(* Logix 5000 project; controller MECO9497 vendor 1 type 14 code 106 rev 21.11; software revision 21.00; part 4 of 4 *)
(* tags used below, declared in another part *)
   AAH_200_SP : REAL;
   AAH_200_SP_H : BOOL;
   AAH_200_SP_N : BOOL;
   AAH_200_SP_O : REAL;
   ALERT_ALARM_SU_DELAY : TIMER;
   ALERT_ALARM_SU_DELAY_H : BOOL;
   ALERT_ALARM_SU_DELAY_N : BOOL;
   ALERT_ALARM_SU_DELAY_O : DINT;
   DIST_COND_ALRM_STARTUP_TIME_H : BOOL;
   DIST_COND_ALRM_STARTUP_TIME_N : BOOL;
   DIST_COND_ALRM_STARTUP_TIME_O : REAL;
   DIST_COND_ALRM_STARTUP_TMR : TIMER;
   DIST_PUMP_START_SP : REAL;
   DIST_PUMP_START_SP_H : BOOL;
   DIST_PUMP_START_SP_N : BOOL;
   DIST_PUMP_START_SP_OIT : REAL;
   DIST_PUMP_STOP_SP : REAL;
   DIST_PUMP_STOP_SP_H : BOOL;
   DIST_PUMP_STOP_SP_N : BOOL;
   DIST_PUMP_STOP_SP_OIT : DINT;
   DSTLT_TEMP_ALRM_SU_DELAY : TIMER;
   DSTLT_TEMP_ALRM_SU_DELAY_H : BOOL;
   DSTLT_TEMP_ALRM_SU_DELAY_N : BOOL;
   DSTLT_TEMP_ALRM_SU_DELAY_O : REAL;
   ENGINEER : BOOL;
   EVAP_PRESSURE_PERM_TIME_H : BOOL;
   EVAP_PRESSURE_PERM_TIME_N : BOOL;
   EVAP_PRESSURE_PERM_TIME_O : REAL;
   EVAP_PRESSURE_PERM_TIMER : TIMER;
   EXCESS_DIST_TIME_SP_H : BOOL;
   EXCESS_DIST_TIME_SP_N : BOOL;
   EXCESS_DIST_TIME_SP_OIT : REAL;
   EXCESS_DSTLT_DRAIN_TIMER : TIMER;
   FC_300_SP : DINT;
   FC_300_SP_H : BOOL;
   FC_300_SP_N : BOOL;
   FC_300_SP_O : DINT;
   IAL_100_SP : REAL;
   IAL_100_SP_H : BOOL;
   IAL_100_SP_N : BOOL;
   IAL_100_SP_OIT : REAL;
   LAAH_100_ALERT_H : BOOL;
   LAAH_100_ALERT_N : BOOL;
   LAAH_100_ALERT_O : DINT;
   LAAH_100_SP : DINT;
   LAAL_100_ALERT_H : BOOL;
   LAAL_100_ALERT_N : BOOL;
   LAAL_100_ALERT_O : DINT;
   LAAL_100_SP : DINT;
   LAH_100_SP : REAL;
   LAH_100_SP_H : BOOL;
   LAH_100_SP_N : BOOL;
   LAH_100_SP_OIT : REAL;
   LAL_100_SP : REAL;
   LAL_100_SP_H : BOOL;
   LAL_100_SP_N : BOOL;
   LAL_100_SP_OIT : REAL;
   LCV_100_AO : ALIAS FOR Local:5:O.Ch2Data;
   LCV_200_AO : ALIAS FOR Local:5:O.Ch3Data;
   LIC_100 : PID;
   LIC_200 : PID;
   LT_100_AI : ALIAS FOR Local:3:I.Ch3Data;
   LT_200_AI : ALIAS FOR Local:3:I.Ch4Data;
   PAAH_103_ALERT_H : BOOL;
   PAAH_103_ALERT_N : BOOL;
   PAAH_103_ALERT_O : REAL;
   PAAH_103_SP : REAL;
   PAAL_103_ALERT_H : BOOL;
   PAAL_103_ALERT_N : BOOL;
   PAAL_103_ALERT_O : REAL;
   PAAL_103_SP : REAL;
   PAH_103_SP : REAL;
   PAH_103_SP_H : BOOL;
   PAH_103_SP_N : BOOL;
   PAH_103_SP_OIT : REAL;
   PAL_103_SP : REAL;
   PAL_103_SP_H : BOOL;
   PAL_103_SP_N : BOOL;
   PAL_103_SP_OIT : REAL;
   PCV_103_AO : ALIAS FOR Local:5:O.Ch0Data;
   PIC_103 : PID;
   PT_103_AI : ALIAS FOR Local:3:I.Ch0Data;
   TAL_200_SP : REAL;
   TAL_200_SP_H : BOOL;
   TAL_200_SP_N : BOOL;
   TAL_200_SP_OIT : REAL;
   TCV_102_AO : ALIAS FOR Local:5:O.Ch4Data;
   TCV_200_AO : ALIAS FOR Local:5:O.Ch1Data;
   TIC_102 : PID;
   TIC_102_CV_SU_H : BOOL;
   TIC_102_CV_SU_N : BOOL;
   TIC_102_CV_SU_O : DINT;
   TIC_102_CV_SU_TIMER : TIMER;
   TIC_200 : PID;
   TT_102_AI : ALIAS FOR Local:3:I.Ch1Data;
   TT_200_AI : ALIAS FOR Local:4:I.Ch1Data;
(* MainProgram, continued *)

ROUTINE SETPOINTS   (* ladder *)
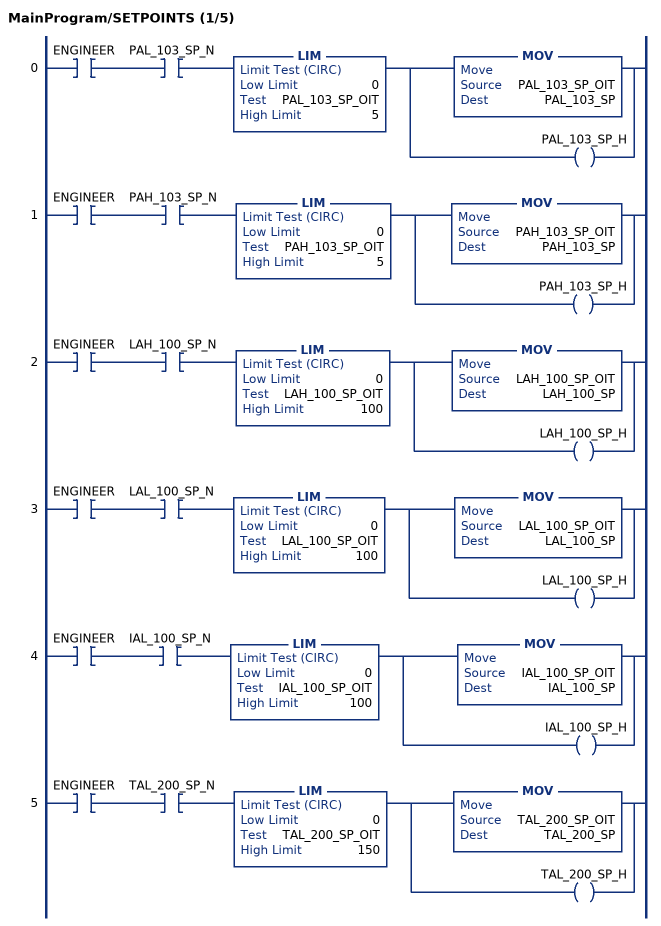
   0: XIC(ENGINEER)XIC(PAL_103_SP_N)LIM(0,PAL_103_SP_OIT,5)[MOV(PAL_103_SP_OIT,PAL_103_SP) ,OTE(PAL_103_SP_H) ];
   1: XIC(ENGINEER)XIC(PAH_103_SP_N)LIM(0,PAH_103_SP_OIT,5)[MOV(PAH_103_SP_OIT,PAH_103_SP) ,OTE(PAH_103_SP_H) ];
   2: XIC(ENGINEER)XIC(LAH_100_SP_N)LIM(0,LAH_100_SP_OIT,100)[MOV(LAH_100_SP_OIT,LAH_100_SP) ,OTE(LAH_100_SP_H) ];
   3: XIC(ENGINEER)XIC(LAL_100_SP_N)LIM(0,LAL_100_SP_OIT,100)[MOV(LAL_100_SP_OIT,LAL_100_SP) ,OTE(LAL_100_SP_H) ];
   4: XIC(ENGINEER)XIC(IAL_100_SP_N)LIM(0,IAL_100_SP_OIT,100)[MOV(IAL_100_SP_OIT,IAL_100_SP) ,OTE(IAL_100_SP_H) ];
   5: XIC(ENGINEER)XIC(TAL_200_SP_N)LIM(0,TAL_200_SP_OIT,150)[MOV(TAL_200_SP_OIT,TAL_200_SP) ,OTE(TAL_200_SP_H) ];
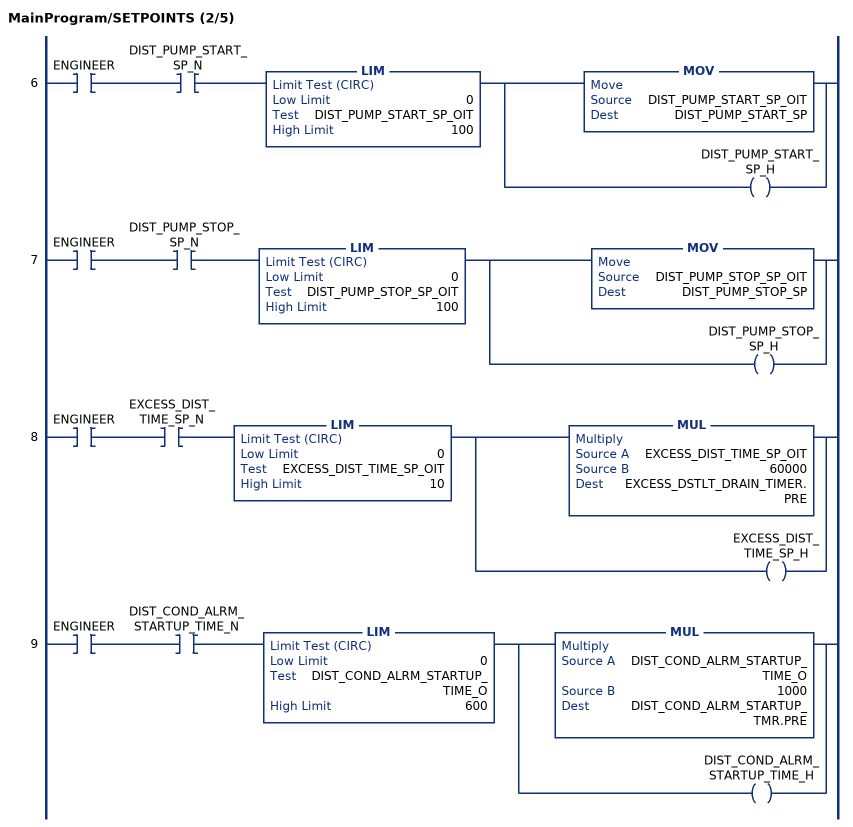
   6: XIC(ENGINEER)XIC(DIST_PUMP_START_SP_N)LIM(0,DIST_PUMP_START_SP_OIT,100)[MOV(DIST_PUMP_START_SP_OIT,DIST_PUMP_START_SP) ,OTE(DIST_PUMP_START_SP_H) ];
   7: XIC(ENGINEER)XIC(DIST_PUMP_STOP_SP_N)LIM(0,DIST_PUMP_STOP_SP_OIT,100)[MOV(DIST_PUMP_STOP_SP_OIT,DIST_PUMP_STOP_SP) ,OTE(DIST_PUMP_STOP_SP_H) ];
   8: XIC(ENGINEER)XIC(EXCESS_DIST_TIME_SP_N)LIM(0,EXCESS_DIST_TIME_SP_OIT,10)[MUL(EXCESS_DIST_TIME_SP_OIT,60000,EXCESS_DSTLT_DRAIN_TIMER.PRE) ,OTE(EXCESS_DIST_TIME_SP_H) ];
   9: XIC(ENGINEER)XIC(DIST_COND_ALRM_STARTUP_TIME_N)LIM(0,DIST_COND_ALRM_STARTUP_TIME_O,600)[MUL(DIST_COND_ALRM_STARTUP_TIME_O,1000,DIST_COND_ALRM_STARTUP_TMR.PRE) ,OTE(DIST_COND_ALRM_STARTUP_TIME_H) ];
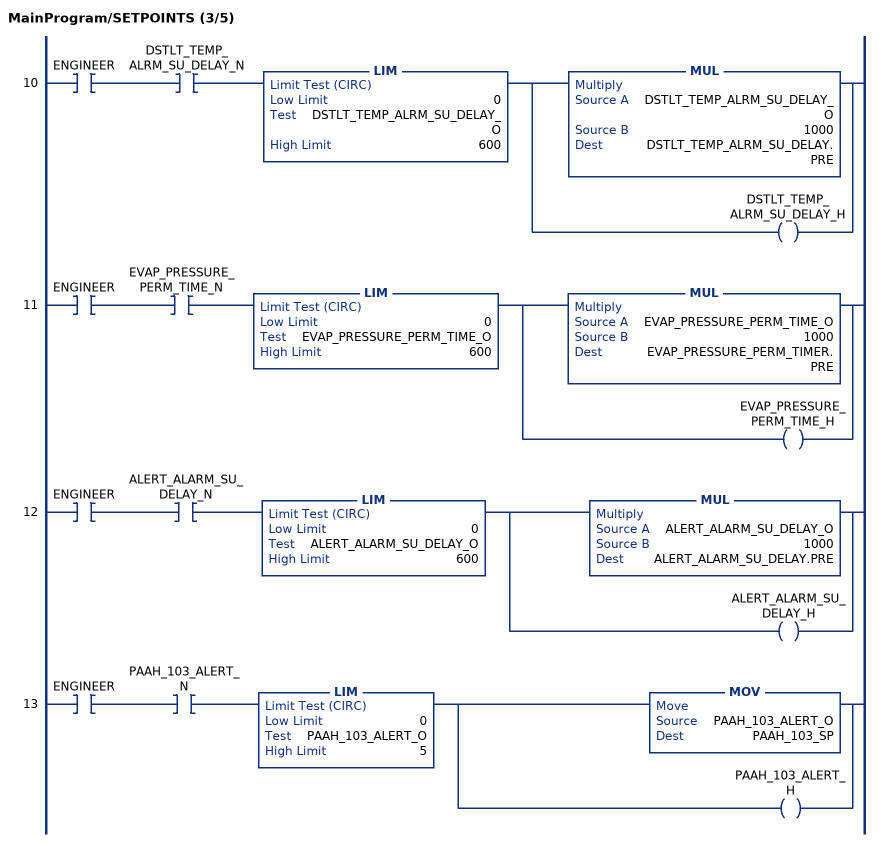
   10: XIC(ENGINEER)XIC(DSTLT_TEMP_ALRM_SU_DELAY_N)LIM(0,DSTLT_TEMP_ALRM_SU_DELAY_O,600)[MUL(DSTLT_TEMP_ALRM_SU_DELAY_O,1000,DSTLT_TEMP_ALRM_SU_DELAY.PRE) ,OTE(DSTLT_TEMP_ALRM_SU_DELAY_H) ];
   11: XIC(ENGINEER)XIC(EVAP_PRESSURE_PERM_TIME_N)LIM(0,EVAP_PRESSURE_PERM_TIME_O,600)[MUL(EVAP_PRESSURE_PERM_TIME_O,1000,EVAP_PRESSURE_PERM_TIMER.PRE) ,OTE(EVAP_PRESSURE_PERM_TIME_H) ];
   12: XIC(ENGINEER)XIC(ALERT_ALARM_SU_DELAY_N)LIM(0,ALERT_ALARM_SU_DELAY_O,600)[MUL(ALERT_ALARM_SU_DELAY_O,1000,ALERT_ALARM_SU_DELAY.PRE) ,OTE(ALERT_ALARM_SU_DELAY_H) ];
   13: XIC(ENGINEER)XIC(PAAH_103_ALERT_N)LIM(0,PAAH_103_ALERT_O,5)[MOV(PAAH_103_ALERT_O,PAAH_103_SP) ,OTE(PAAH_103_ALERT_H) ];
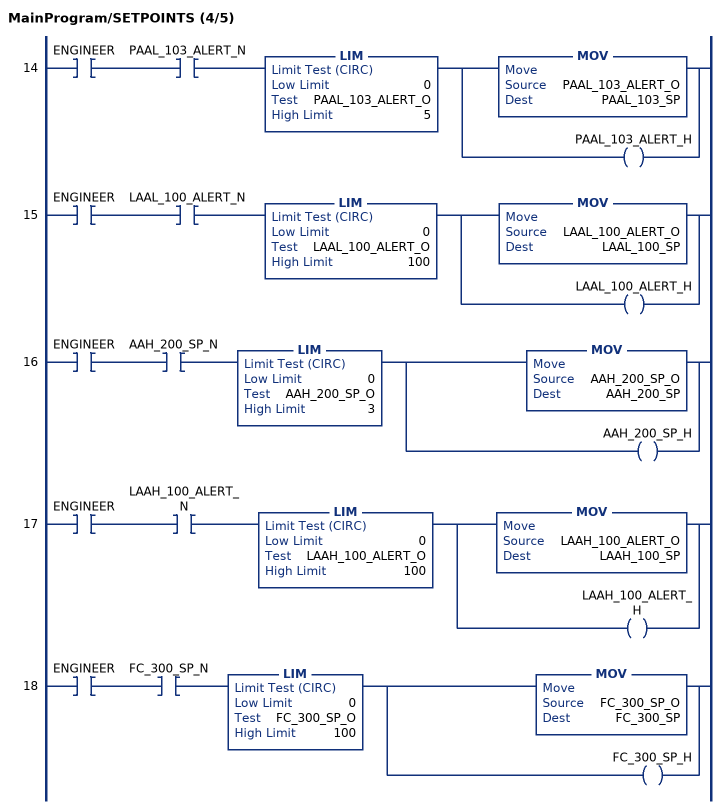
   14: XIC(ENGINEER)XIC(PAAL_103_ALERT_N)LIM(0,PAAL_103_ALERT_O,5)[MOV(PAAL_103_ALERT_O,PAAL_103_SP) ,OTE(PAAL_103_ALERT_H) ];
   15: XIC(ENGINEER)XIC(LAAL_100_ALERT_N)LIM(0,LAAL_100_ALERT_O,100)[MOV(LAAL_100_ALERT_O,LAAL_100_SP) ,OTE(LAAL_100_ALERT_H) ];
   16: XIC(ENGINEER)XIC(AAH_200_SP_N)LIM(0,AAH_200_SP_O,3)[MOV(AAH_200_SP_O,AAH_200_SP) ,OTE(AAH_200_SP_H) ];
   17: XIC(ENGINEER)XIC(LAAH_100_ALERT_N)LIM(0,LAAH_100_ALERT_O,100)[MOV(LAAH_100_ALERT_O,LAAH_100_SP) ,OTE(LAAH_100_ALERT_H) ];
   18: XIC(ENGINEER)XIC(FC_300_SP_N)LIM(0,FC_300_SP_O,100)[MOV(FC_300_SP_O,FC_300_SP) ,OTE(FC_300_SP_H) ];
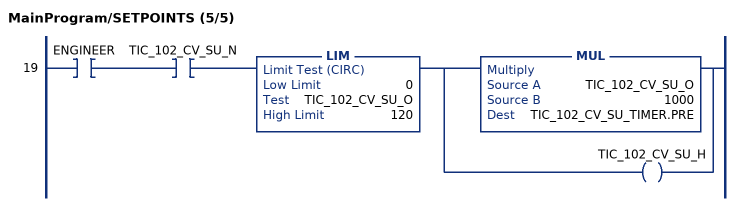
   19: XIC(ENGINEER)XIC(TIC_102_CV_SU_N)LIM(0,TIC_102_CV_SU_O,120)[MUL(TIC_102_CV_SU_O,1000,TIC_102_CV_SU_TIMER.PRE) ,OTE(TIC_102_CV_SU_H) ];
END_ROUTINE
END_PROGRAM

PROGRAM PID_MAIN   (* main routine PID_MIAN_ROUTINE *)

ROUTINE PID_MIAN_ROUTINE   (* ladder *)
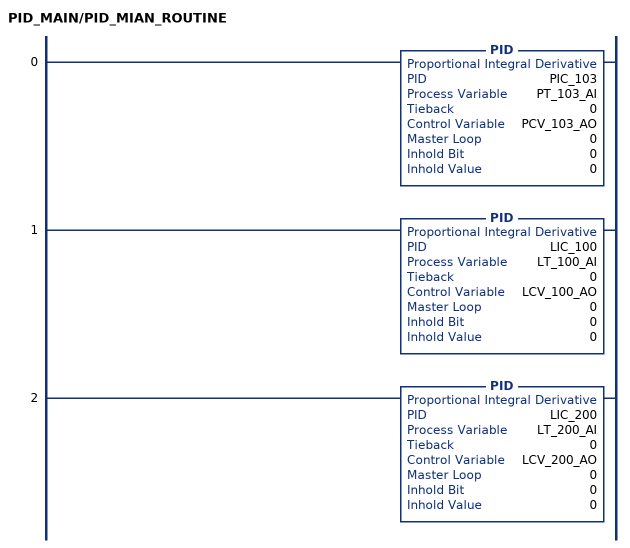
   0: PID(PIC_103,PT_103_AI,0,PCV_103_AO,0,0,0);
   1: PID(LIC_100,LT_100_AI,0,LCV_100_AO,0,0,0);
   2: PID(LIC_200,LT_200_AI,0,LCV_200_AO,0,0,0);
END_ROUTINE
END_PROGRAM

PROGRAM PID_SLOW   (* main routine PID_SLOW_ROUTINE *)

ROUTINE PID_SLOW_ROUTINE   (* ladder *)
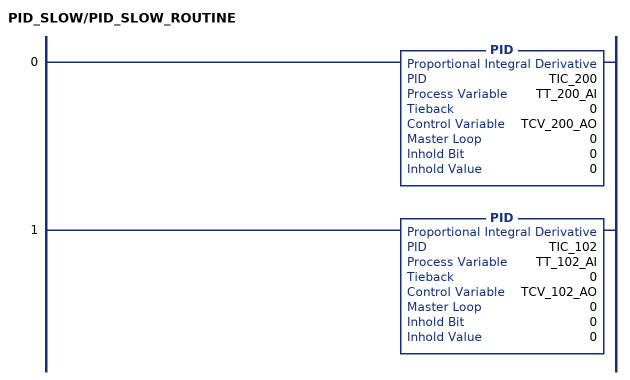
   0: PID(TIC_200,TT_200_AI,0,TCV_200_AO,0,0,0);
   1: PID(TIC_102,TT_102_AI,0,TCV_102_AO,0,0,0);
END_ROUTINE
END_PROGRAM
